Fanuc KAREL source: KT00516.KL

PROGRAM KT00516
%NOLOCKGROUP
VAR
  P1: XYZWPREXT
  P2: POSITION
  OUT: XYZWPREXT
BEGIN
  P1.X = 1.0
  OUT = P1 : P2
END KT00516
